Omron CX-Programmer project NewProject (CX-Programmer 9.75)

# PLC robotBox: CP1E N30

## Global symbols (name address type ; comment)
0.00 BOOL  ; f5
0.01 BOOL  ; x0
0.02 BOOL  ; x1
0.03 BOOL  ; x2
0.04 BOOL  ; x3
0.05 BOOL  ; S reset
100.00 BOOL  ; robot
100.01 BOOL  ; konveyor
100.02 BOOL  ; Upper
100.03 BOOL  ; Middle
100.04 BOOL  ; Lower

## Program NewProgram1 (cyclic task 0)

### Section Section1

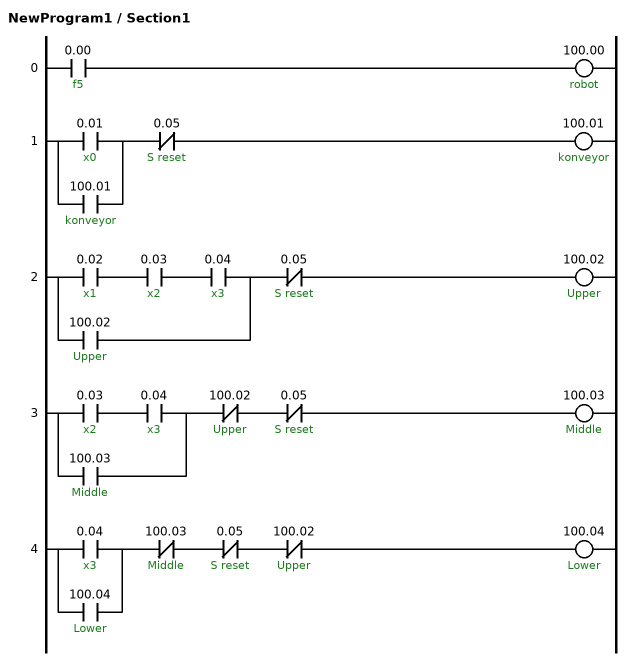
; rung 0
LD 0.00  ; f5
OUT 100.00  ; robot
; rung 1
LD 0.01  ; x0
OR 100.01  ; konveyor
ANDNOT 0.05  ; S reset
OUT 100.01  ; konveyor
; rung 2
LD 0.02  ; x1
AND 0.03  ; x2
AND 0.04  ; x3
OR 100.02  ; Upper
ANDNOT 0.05  ; S reset
OUT 100.02  ; Upper
; rung 3
LD 0.03  ; x2
AND 0.04  ; x3
OR 100.03  ; Middle
ANDNOT 100.02  ; Upper
ANDNOT 0.05  ; S reset
OUT 100.03  ; Middle
; rung 4
LD 0.04  ; x3
OR 100.04  ; Lower
ANDNOT 100.03  ; Middle
ANDNOT 0.05  ; S reset
ANDNOT 100.02  ; Upper
OUT 100.04  ; Lower

### Section END
; rung 0
END(001)